FUNCTION_BLOCK PUBLIC FB_Piston_U_L// EXTENDS FB_Piston
VAR_INPUT
	enable		: BOOL	;
	sen_Upper	: BOOL	;
	sen_Lower	: BOOL	;

END_VAR
VAR_OUTPUT
	valve_Upper		:BOOL;
	valve_Lower		:BOOL;	
END_VAR
VAR
	tOn: TIME:=T#1S;
	tOff: TIME:=T#1S;
	Call_RTrig_ReqUp: R_TRIG;
	Call_RTrig_ReqLow: R_TRIG;
	
	b_Memo_ReqUp	:	BOOL	;
	b_Memo_ReqLow	:	BOOL	;
	Call_FTrig_Error: 	F_TRIG	;
	stPis			:	REFERENCE TO ST_Piston;
	ton_req_Upper: TON;
	ton_req_Lower: TON;
	tOperation: TIME := T#2S;
	ton_err_Upper: TON;
	ton_err_Lower: TON;
	tError: TIME := T#5s;
END_VAR
VAR_IN_OUT
	st_Piston_U_L	:	ST_Piston_U_L	;
	stOperation		: ST_OperationButtons;
END_VAR

act_Get_Reference();
act_SetOutputs();

IF stPis.b_Error THEN;
	stOperation.bSetPause:=TRUE;
END_IF

ton_req_Upper(PT:=tOperation, IN:=st_Piston_U_L.req_Upper);
ton_req_Lower(PT:=tOperation, IN:=st_Piston_U_L.req_Lower);

ton_err_Upper(PT:=tError);
ton_err_Lower(PT:=tError);

IF TRUE 
AND st_Piston_U_L.req_Upper
AND (NOT st_Piston_U_L.st_Upper)
AND (NOT FALSE) // reset error
THEN;
	ton_err_Upper.IN:=TRUE;
ELSE;
	ton_err_Upper.IN:=FALSE;
END_IF

IF TRUE 
AND st_Piston_U_L.req_Lower
AND (NOT st_Piston_U_L.st_Lower)
AND (NOT FALSE) // reset error
THEN;
	ton_err_Lower.IN:=TRUE;
ELSE;
	ton_err_Lower.IN:=FALSE;
END_IF

IF ton_err_Upper.Q OR ton_err_Lower.Q THEN;
	stPis.b_Error:=TRUE;
END_IF

ACTION act_Get_Reference:
//st_Piston_U_L.str_Piston REF= g_Piston.stPis[iFB_Num];
stPis REF= g_Piston.stPis[st_Piston_U_L.iFB_Num];
END_ACTION

ACTION act_SetOutputs:
(*IF st_Piston_U_L.bError THEN
	IF st_Piston_U_L.req_Upper THEN
		b_Memo_ReqUp:=TRUE;
	END_IF
	IF st_Piston_U_L.req_Lower THEN
		b_Memo_ReqLow:=TRUE;
	END_IF
	st_Piston_U_L.req_Upper:=FALSE;
	st_Piston_U_L.req_Lower:=FALSE;
END_IF*)

(*
Call_FTrig_Error(CLK:=st_Piston_U_L.bError , Q=> );

IF Call_FTrig_Error.Q THEN
	st_Piston_U_L.req_Upper:=b_Memo_ReqUp;
	st_Piston_U_L.req_Lower:=b_Memo_ReqLow;
	b_Memo_ReqUp:=FALSE;
	b_Memo_ReqLow:=FALSE;
END_IF*)

//Resseting opposite signal
//***************************************************************
Call_RTrig_ReqUp(CLK:=st_Piston_U_L.req_Upper , Q=> );
Call_RTrig_ReqLow(CLK:=st_Piston_U_L.req_Lower, Q=> );
IF Call_RTrig_ReqUp.Q THEN
	st_Piston_U_L.req_Lower:=FALSE;
END_IF

IF Call_RTrig_ReqLow.Q THEN
	st_Piston_U_L.req_Upper :=FALSE;
END_IF
//***************************************************************

IF enable AND stPis.valve_Close THEN;
	st_Piston_U_L.exist:=TRUE;
	
	IF st_Piston_U_L.req_Upper THEN;
		valve_Upper:=TRUE;
		valve_Lower:=FALSE;		
	ELSIF st_Piston_U_L.req_Lower THEN;
		valve_Upper:=FALSE;
		valve_Lower:=TRUE;		
	ELSE;
		valve_Upper:=FALSE;
		valve_Lower:=FALSE;		
	END_IF
ELSE;
	st_Piston_U_L.exist:=FALSE;
	st_Piston_U_L.req_Upper:=FALSE;
	st_Piston_U_L.req_Lower:=FALSE;
	valve_Upper:=FALSE;
	valve_Lower:=FALSE;
END_IF

//outputs for hmi
st_Piston_U_L.out_Upper:=valve_Upper;
st_Piston_U_L.out_Lower:=valve_Lower;

//Status
st_Piston_U_L.st_Upper:=m_sen_Upper();
st_Piston_U_L.st_Lower:=m_sen_Lower();
st_Piston_U_L.st_Released:=(NOT m_sen_Upper() AND NOT m_sen_Lower());

st_Piston_U_L.sen_Upper:=sen_Upper;
st_Piston_U_L.sen_Lower:=sen_Lower;
END_ACTION

METHOD m_sen_Lower : BOOL
VAR_INPUT
END_VAR
IF st_Piston_U_L.sen_Lower_exist THEN; // sensor exist
	m_sen_Lower:=sen_Lower;
ELSE;
	m_sen_Lower:=ton_req_Lower.Q;
END_IF
END_METHOD

METHOD m_sen_Upper : BOOL
VAR_INPUT
END_VAR
IF st_Piston_U_L.sen_Upper_exist THEN; // sensor exist
	m_sen_Upper:=sen_Upper;
ELSE;
	m_sen_Upper:=ton_req_Upper.Q;
END_IF
END_METHOD

END_FUNCTION_BLOCK

(* stored: Version 1.1.0.1, ProductVersion 3.1.4024.13
   POU FB_Piston_U_L: Id {f6df062b-8dd7-4dca-98fe-56ea9e281485}, SpecialFunc None
   Action act_Get_Reference: Id {60607663-ce4f-44c4-8288-4340f34ed98c}
   Action act_SetOutputs: Id {fe9d830e-c8cb-470f-9da2-a61c532c4f0f}
   Method m_sen_Lower: Id {87f5513f-eed4-4f44-8483-3e0613ae32b6}
   Method m_sen_Upper: Id {2404f77a-a933-4805-88d7-69cc1f20bd1a} *)
